DATA_BLOCK "GDB_AlarmPersistTest"
{ S7_Optimized_Access := 'TRUE' }
VERSION : 0.1
NON_RETAIN
VAR
    Operation : Int;
    UnicodeMode : Int;
    Scope : String[80];
    Text : WString[255];
    Reason : DInt;
    Slot {ExternalWritable := 'False'} : Int;
    Generation {ExternalWritable := 'False'} : UDInt;
    Checksum {ExternalWritable := 'False'} : DWord;
    Used {ExternalWritable := 'False'} : Int;
    Applied {ExternalWritable := 'False'} : Bool;
END_VAR
BEGIN
END_DATA_BLOCK
